(* IEC 61131-3 sources: plc-st-coding-agent/progress/evidence/f14_v3_parallel_20261112/jobs/custom_deepseek-v4pro (part 3) *)

(* ---- self-hard-07.raw_candidate_01.st ---- *)
FUNCTION_BLOCK FB
VAR_INPUT
    mode : INT;
    resetBtn : BOOL;
    scanSeconds : REAL;
    tempSP : REAL;
    tempPV : REAL;
    flowPV : REAL;
    manualFlowSP : REAL;
    manualValve : REAL;
END_VAR
VAR_OUTPUT
    flowSP : REAL;
    valveCommand : REAL;
    fault : BOOL;
    normalMode : BOOL;
END_VAR
VAR
    hasPrev : BOOL := FALSE;
    prevMode : INT := 0;
    prevReset : BOOL := FALSE;
    prevFlowSP : REAL := 0.0;
    prevValveCommand : REAL := 0.0;
    prevET : REAL := 0.0;
    prevEF : REAL := 0.0;
    resetRising : BOOL;
    eT : REAL;
    eF : REAL;
    flowRaw : REAL;
    valveRaw : REAL;
    trialT : REAL;
    trialF : REAL;
END_VAR

fault := (mode < 0) OR (mode > 2) OR (scanSeconds <= 0.0) OR (scanSeconds > 10.0);
resetRising := resetBtn AND NOT prevReset;

IF NOT hasPrev THEN
    normalMode := FALSE;
    flowSP := manualFlowSP;
    valveCommand := manualValve;
ELSIF resetRising THEN
    normalMode := FALSE;
    flowSP := manualFlowSP;
    valveCommand := manualValve;
ELSIF fault THEN
    normalMode := FALSE;
    flowSP := manualFlowSP;
    valveCommand := manualValve;
ELSIF mode <> prevMode THEN
    normalMode := FALSE;
    IF mode = 2 THEN
        flowSP := prevFlowSP;
        valveCommand := prevValveCommand;
    ELSE
        flowSP := manualFlowSP;
        valveCommand := prevValveCommand;
    END_IF;
ELSE
    normalMode := TRUE;
    IF mode = 0 THEN
        flowSP := manualFlowSP;
        valveCommand := manualValve;
    ELSIF mode = 1 THEN
        flowSP := manualFlowSP;
        eF := flowSP - flowPV;
        trialF := prevValveCommand - 2.0 * prevEF + 0.5 * eF * scanSeconds;
        valveRaw := 2.0 * eF + trialF;
        valveCommand := LIMIT(0.0, valveRaw, 100.0);
    ELSIF mode = 2 THEN
        eT := tempSP - tempPV;
        trialT := prevFlowSP - 1.0 * prevET + 0.2 * eT * scanSeconds;
        flowRaw := 1.0 * eT + trialT;
        flowSP := LIMIT(0.0, flowRaw, 50.0);
        eF := flowSP - flowPV;
        trialF := prevValveCommand - 2.0 * prevEF + 0.5 * eF * scanSeconds;
        valveRaw := 2.0 * eF + trialF;
        valveCommand := LIMIT(0.0, valveRaw, 100.0);
    END_IF;
END_IF;

prevFlowSP := flowSP;
prevValveCommand := valveCommand;
prevET := tempSP - tempPV;
prevEF := flowSP - flowPV;
prevMode := mode;
prevReset := resetBtn;
hasPrev := TRUE;

END_FUNCTION_BLOCK

(* ---- self-medium-01.candidate_01.st ---- *)
FUNCTION_BLOCK FB
VAR_INPUT
    recipe : ARRAY[1..8] OF ST_Recipe;   // 配方槽位 1..8，槽位 recipeID=0 表示空
    selSlot : INT;                        // 操作员选中的槽位，合法范围 1..8
    loadCmd : BOOL;                       // 装载命令（上升沿触发一次装载）
    running : BOOL;                       // 当前是否处于生产状态
END_VAR
VAR_OUTPUT
    valid : BOOL;                         // 配方校验通过
    loadedID : INT;                       // 已装载的配方号，无配方时为 0
END_VAR
VAR
    prevLoadCmd  : BOOL;                  // 上一扫描周期的 loadCmd
    prevValid    : BOOL;                  // 上一扫描周期的 valid 输出
    prevLoadedID : INT;                   // 上一扫描周期的 loadedID 输出
    edge         : BOOL;                  // loadCmd 上升沿标志
    slotIndex    : INT;                   // 合法的槽位下标
    slotRecipe   : ST_Recipe;             // 当前选中的配方结构体
    ratioOK      : BOOL;                  // totalRatio 是否在合法区间
    tempOK       : BOOL;                  // temperature 是否在合法区间
END_VAR

    // 计算装载命令的上升沿
    edge := loadCmd AND NOT prevLoadCmd;

    IF running THEN
        // 生产状态：保持上一拍输出，包括刚进入生产的第一拍
        valid := prevValid;
        loadedID := prevLoadedID;
    ELSIF edge THEN
        // 非生产状态且检测到装载命令上升沿
        // 检查槽位是否越界
        IF (selSlot < 1) OR (selSlot > 8) THEN
            // 越界：判为非法，且不得访问数组外内存
            valid := FALSE;
            loadedID := 0;
        ELSE
            // 合法槽位
            slotIndex := selSlot;
            slotRecipe := recipe[slotIndex];

            // 检查槽位是否为空
            IF slotRecipe.recipeID = 0 THEN
                // 空槽：非法
                valid := FALSE;
                loadedID := 0;
            ELSE
                // 检查总配比和温度
                ratioOK := (slotRecipe.totalRatio >= 99.0) AND (slotRecipe.totalRatio <= 101.0);
                tempOK  := (slotRecipe.temperature >= 30.0) AND (slotRecipe.temperature <= 180.0);

                IF ratioOK AND tempOK THEN
                    // 全部校验通过
                    valid := TRUE;
                    loadedID := slotRecipe.recipeID;
                ELSE
                    // 任一校验失败
                    valid := FALSE;
                    loadedID := 0;
                END_IF;
            END_IF;
        END_IF;
    ELSE
        // 无装载沿且未生产：保持上一拍输出
        valid := prevValid;
        loadedID := prevLoadedID;
    END_IF;

    // 更新历史状态
    prevLoadCmd  := loadCmd;
    prevValid    := valid;
    prevLoadedID := loadedID;
END_FUNCTION_BLOCK

(* ---- self-medium-01.candidate_02.st ---- *)
TYPE ST_Recipe :
STRUCT
    recipeID : INT;
    totalRatio : REAL;
    temperature : REAL;
END_STRUCT;
END_TYPE;

FUNCTION_BLOCK FB
VAR_INPUT
    recipe : ARRAY[1..8] OF ST_Recipe;
    selSlot : INT;
    loadCmd : BOOL;
    running : BOOL;
END_VAR
VAR_OUTPUT
    valid : BOOL;
    loadedID : INT;
END_VAR
VAR
    prevLoadCmd  : BOOL;
    prevValid    : BOOL;
    prevLoadedID : INT;
    edge         : BOOL;
    slotIndex    : INT;
    slotRecipe   : ST_Recipe;
    ratioOK      : BOOL;
    tempOK       : BOOL;
END_VAR

    edge := loadCmd AND NOT prevLoadCmd;

    IF running THEN
        (* 生产状态：保持上一拍输出，包括刚进入生产的第一拍 *)
        valid := prevValid;
        loadedID := prevLoadedID;
    ELSIF edge THEN
        (* 非生产状态且检测到装载命令上升沿 *)
        IF (selSlot < 1) OR (selSlot > 8) THEN
            (* 槽位越界：判为非法，不访问数组 *)
            valid := FALSE;
            loadedID := 0;
        ELSE
            slotIndex := selSlot;
            slotRecipe := recipe[slotIndex];

            IF slotRecipe.recipeID = 0 THEN
                (* 空槽：非法 *)
                valid := FALSE;
                loadedID := 0;
            ELSE
                ratioOK := (slotRecipe.totalRatio >= 99.0) AND (slotRecipe.totalRatio <= 101.0);
                tempOK  := (slotRecipe.temperature >= 30.0) AND (slotRecipe.temperature <= 180.0);

                IF ratioOK AND tempOK THEN
                    valid := TRUE;
                    loadedID := slotRecipe.recipeID;
                ELSE
                    valid := FALSE;
                    loadedID := 0;
                END_IF;
            END_IF;
        END_IF;
    ELSE
        (* 无装载沿且未生产：保持上一拍输出 *)
        valid := prevValid;
        loadedID := prevLoadedID;
    END_IF;

    (* 更新历史状态 *)
    prevLoadCmd  := loadCmd;
    prevValid    := valid;
    prevLoadedID := loadedID;
END_FUNCTION_BLOCK

(* ---- self-medium-01.raw_candidate_01.st ---- *)
FUNCTION_BLOCK FB
VAR_INPUT
    recipe : ARRAY[1..8] OF ST_Recipe;   // 配方槽位 1..8，槽位 recipeID=0 表示空
    selSlot : INT;                        // 操作员选中的槽位，合法范围 1..8
    loadCmd : BOOL;                       // 装载命令（上升沿触发一次装载）
    running : BOOL;                       // 当前是否处于生产状态
END_VAR
VAR_OUTPUT
    valid : BOOL;                         // 配方校验通过
    loadedID : INT;                       // 已装载的配方号，无配方时为 0
END_VAR
VAR
    prevLoadCmd  : BOOL;                  // 上一扫描周期的 loadCmd
    prevValid    : BOOL;                  // 上一扫描周期的 valid 输出
    prevLoadedID : INT;                   // 上一扫描周期的 loadedID 输出
    edge         : BOOL;                  // loadCmd 上升沿标志
    slotIndex    : INT;                   // 合法的槽位下标
    slotRecipe   : ST_Recipe;             // 当前选中的配方结构体
    ratioOK      : BOOL;                  // totalRatio 是否在合法区间
    tempOK       : BOOL;                  // temperature 是否在合法区间
END_VAR

    // 计算装载命令的上升沿
    edge := loadCmd AND NOT prevLoadCmd;

    IF running THEN
        // 生产状态：保持上一拍输出，包括刚进入生产的第一拍
        valid := prevValid;
        loadedID := prevLoadedID;
    ELSIF edge THEN
        // 非生产状态且检测到装载命令上升沿
        // 检查槽位是否越界
        IF (selSlot < 1) OR (selSlot > 8) THEN
            // 越界：判为非法，且不得访问数组外内存
            valid := FALSE;
            loadedID := 0;
        ELSE
            // 合法槽位
            slotIndex := selSlot;
            slotRecipe := recipe[slotIndex];

            // 检查槽位是否为空
            IF slotRecipe.recipeID = 0 THEN
                // 空槽：非法
                valid := FALSE;
                loadedID := 0;
            ELSE
                // 检查总配比和温度
                ratioOK := (slotRecipe.totalRatio >= 99.0) AND (slotRecipe.totalRatio <= 101.0);
                tempOK  := (slotRecipe.temperature >= 30.0) AND (slotRecipe.temperature <= 180.0);

                IF ratioOK AND tempOK THEN
                    // 全部校验通过
                    valid := TRUE;
                    loadedID := slotRecipe.recipeID;
                ELSE
                    // 任一校验失败
                    valid := FALSE;
                    loadedID := 0;
                END_IF;
            END_IF;
        END_IF;
    ELSE
        // 无装载沿且未生产：保持上一拍输出
        valid := prevValid;
        loadedID := prevLoadedID;
    END_IF;

    // 更新历史状态
    prevLoadCmd  := loadCmd;
    prevValid    := valid;
    prevLoadedID := loadedID;
END_FUNCTION_BLOCK

(* ---- self-medium-01.raw_candidate_02.st ---- *)
TYPE ST_Recipe :
STRUCT
    recipeID : INT;
    totalRatio : REAL;
    temperature : REAL;
END_STRUCT
END_TYPE

FUNCTION_BLOCK FB
VAR_INPUT
    recipe : ARRAY[1..8] OF ST_Recipe;
    selSlot : INT;
    loadCmd : BOOL;
    running : BOOL;
END_VAR
VAR_OUTPUT
    valid : BOOL;
    loadedID : INT;
END_VAR
VAR
    prevLoadCmd  : BOOL;
    prevValid    : BOOL;
    prevLoadedID : INT;
    edge         : BOOL;
    slotIndex    : INT;
    slotRecipe   : ST_Recipe;
    ratioOK      : BOOL;
    tempOK       : BOOL;
END_VAR

    edge := loadCmd AND NOT prevLoadCmd;

    IF running THEN
        (* 生产状态：保持上一拍输出，包括刚进入生产的第一拍 *)
        valid := prevValid;
        loadedID := prevLoadedID;
    ELSIF edge THEN
        (* 非生产状态且检测到装载命令上升沿 *)
        IF (selSlot < 1) OR (selSlot > 8) THEN
            (* 槽位越界：判为非法，不访问数组 *)
            valid := FALSE;
            loadedID := 0;
        ELSE
            slotIndex := selSlot;
            slotRecipe := recipe[slotIndex];

            IF slotRecipe.recipeID = 0 THEN
                (* 空槽：非法 *)
                valid := FALSE;
                loadedID := 0;
            ELSE
                ratioOK := (slotRecipe.totalRatio >= 99.0) AND (slotRecipe.totalRatio <= 101.0);
                tempOK  := (slotRecipe.temperature >= 30.0) AND (slotRecipe.temperature <= 180.0);

                IF ratioOK AND tempOK THEN
                    valid := TRUE;
                    loadedID := slotRecipe.recipeID;
                ELSE
                    valid := FALSE;
                    loadedID := 0;
                END_IF;
            END_IF;
        END_IF;
    ELSE
        (* 无装载沿且未生产：保持上一拍输出 *)
        valid := prevValid;
        loadedID := prevLoadedID;
    END_IF;

    (* 更新历史状态 *)
    prevLoadCmd  := loadCmd;
    prevValid    := valid;
    prevLoadedID := loadedID;
END_FUNCTION_BLOCK

(* ---- self-medium-02.candidate_01.st ---- *)
FUNCTION_BLOCK FB
VAR_INPUT
    enable : BOOL;
    rawValue : REAL;
END_VAR
VAR_OUTPUT
    filteredValue : REAL;
    windowFull : BOOL;
    sampleCount : INT;
END_VAR
VAR
    buffer : ARRAY[0..7] OF REAL;
    bufIdx : INT := 0;
    cnt : INT := 0;
    sum : REAL;
    i : INT;
END_VAR

IF enable THEN
    buffer[bufIdx] := rawValue;
    bufIdx := bufIdx + 1;
    IF bufIdx >= 8 THEN
        bufIdx := 0;
    END_IF;

    IF cnt < 8 THEN
        cnt := cnt + 1;
    END_IF;

    sum := 0.0;
    FOR i := 0 TO cnt - 1 DO
        sum := sum + buffer[i];
    END_FOR;

    filteredValue := sum / INT_TO_REAL(cnt);
    sampleCount := cnt;
    windowFull := (cnt >= 8);
ELSE
    cnt := 0;
    bufIdx := 0;
    sampleCount := 0;
    windowFull := FALSE;
END_IF;

END_FUNCTION_BLOCK

(* ---- self-medium-02.raw_candidate_01.st ---- *)
FUNCTION_BLOCK FB
VAR_INPUT
    enable : BOOL;
    rawValue : REAL;
END_VAR
VAR_OUTPUT
    filteredValue : REAL;
    windowFull : BOOL;
    sampleCount : INT;
END_VAR
VAR
    buffer : ARRAY[0..7] OF REAL;
    bufIdx : INT := 0;
    cnt : INT := 0;
    sum : REAL;
    i : INT;
END_VAR

IF enable THEN
    buffer[bufIdx] := rawValue;
    bufIdx := bufIdx + 1;
    IF bufIdx >= 8 THEN
        bufIdx := 0;
    END_IF;

    IF cnt < 8 THEN
        cnt := cnt + 1;
    END_IF;

    sum := 0.0;
    FOR i := 0 TO cnt - 1 DO
        sum := sum + buffer[i];
    END_FOR;

    filteredValue := sum / INT_TO_REAL(cnt);
    sampleCount := cnt;
    windowFull := (cnt >= 8);
ELSE
    cnt := 0;
    bufIdx := 0;
    sampleCount := 0;
    windowFull := FALSE;
END_IF;

END_FUNCTION_BLOCK

(* ---- self-medium-03.candidate_01.st ---- *)
FUNCTION_BLOCK FB
VAR_INPUT
    openBtn : BOOL;
    closeBtn : BOOL;
    openLimit : BOOL;
    closeLimit : BOOL;
    obstacle : BOOL;
END_VAR
VAR_OUTPUT
    motorUp : BOOL;
    motorDown : BOOL;
    errorFlag : BOOL;
END_VAR
VAR
    state : INT := 0; (* 0=IDLE, 1=OPENING, 2=CLOSING, 3=FAULT *)
    preOpenBtn : BOOL := FALSE;
    preCloseBtn : BOOL := FALSE;
    risingOpen : BOOL;
    risingClose : BOOL;
    combo : BOOL;
    preCombo : BOOL;
    risingCombo : BOOL;
END_VAR

(* 计算上升沿 *)
risingOpen := openBtn AND NOT preOpenBtn;
risingClose := closeBtn AND NOT preCloseBtn;
combo := openBtn AND closeBtn;
preCombo := preOpenBtn AND preCloseBtn;
risingCombo := combo AND NOT preCombo;

IF obstacle THEN
    (* 障碍优先：任何状态立即停机并置故障 *)
    state := 3;
    motorUp := FALSE;
    motorDown := FALSE;
    errorFlag := TRUE;
ELSE
    IF state = 3 THEN
        (* 无障碍时的故障处理 *)
        IF risingCombo THEN
            (* 双键组合新上升沿：人工复位 *)
            state := 0;
            motorUp := FALSE;
            motorDown := FALSE;
            errorFlag := FALSE;
        ELSE
            (* 保持故障锁存 *)
            motorUp := FALSE;
            motorDown := FALSE;
            errorFlag := TRUE;
        END_IF;
    ELSE
        (* 非故障状态 *)
        IF (state = 1 AND openLimit) OR (state = 2 AND closeLimit) THEN
            (* 到达本方向限位：停机回IDLE *)
            state := 0;
            motorUp := FALSE;
            motorDown := FALSE;
            errorFlag := FALSE;
        ELSE
            IF state = 1 THEN
                (* 开门运行中 *)
                motorUp := TRUE;
                motorDown := FALSE;
                errorFlag := FALSE;
                (* state 保持 1 *)
            ELSIF state = 2 THEN
                (* 关门运行中 *)
                motorUp := FALSE;
                motorDown := TRUE;
                errorFlag := FALSE;
                (* state 保持 2 *)
            ELSE
                (* IDLE状态 *)
                IF risingOpen AND NOT closeBtn AND NOT openLimit THEN
                    state := 1;
                    motorUp := TRUE;
                    motorDown := FALSE;
                    errorFlag := FALSE;
                ELSIF risingClose AND NOT openBtn AND NOT closeLimit THEN
                    state := 2;
                    motorUp := FALSE;
                    motorDown := TRUE;
                    errorFlag := FALSE;
                ELSE
                    motorUp := FALSE;
                    motorDown := FALSE;
                    errorFlag := FALSE;
                    state := 0; (* 保持IDLE *)
                END_IF;
            END_IF;
        END_IF;
    END_IF;
END_IF;

(* 更新上一拍按钮状态 *)
preOpenBtn := openBtn;
preCloseBtn := closeBtn;

END_FUNCTION_BLOCK

(* ---- self-medium-03.raw_candidate_01.st ---- *)
FUNCTION_BLOCK FB
VAR_INPUT
    openBtn : BOOL;
    closeBtn : BOOL;
    openLimit : BOOL;
    closeLimit : BOOL;
    obstacle : BOOL;
END_VAR
VAR_OUTPUT
    motorUp : BOOL;
    motorDown : BOOL;
    errorFlag : BOOL;
END_VAR
VAR
    state : INT := 0; (* 0=IDLE, 1=OPENING, 2=CLOSING, 3=FAULT *)
    preOpenBtn : BOOL := FALSE;
    preCloseBtn : BOOL := FALSE;
    risingOpen : BOOL;
    risingClose : BOOL;
    combo : BOOL;
    preCombo : BOOL;
    risingCombo : BOOL;
END_VAR

(* 计算上升沿 *)
risingOpen := openBtn AND NOT preOpenBtn;
risingClose := closeBtn AND NOT preCloseBtn;
combo := openBtn AND closeBtn;
preCombo := preOpenBtn AND preCloseBtn;
risingCombo := combo AND NOT preCombo;

IF obstacle THEN
    (* 障碍优先：任何状态立即停机并置故障 *)
    state := 3;
    motorUp := FALSE;
    motorDown := FALSE;
    errorFlag := TRUE;
ELSE
    IF state = 3 THEN
        (* 无障碍时的故障处理 *)
        IF risingCombo THEN
            (* 双键组合新上升沿：人工复位 *)
            state := 0;
            motorUp := FALSE;
            motorDown := FALSE;
            errorFlag := FALSE;
        ELSE
            (* 保持故障锁存 *)
            motorUp := FALSE;
            motorDown := FALSE;
            errorFlag := TRUE;
        END_IF
    ELSE
        (* 非故障状态 *)
        IF (state = 1 AND openLimit) OR (state = 2 AND closeLimit) THEN
            (* 到达本方向限位：停机回IDLE *)
            state := 0;
            motorUp := FALSE;
            motorDown := FALSE;
            errorFlag := FALSE;
        ELSE
            IF state = 1 THEN
                (* 开门运行中 *)
                motorUp := TRUE;
                motorDown := FALSE;
                errorFlag := FALSE;
                (* state 保持 1 *)
            ELSIF state = 2 THEN
                (* 关门运行中 *)
                motorUp := FALSE;
                motorDown := TRUE;
                errorFlag := FALSE;
                (* state 保持 2 *)
            ELSE
                (* IDLE状态 *)
                IF risingOpen AND NOT closeBtn AND NOT openLimit THEN
                    state := 1;
                    motorUp := TRUE;
                    motorDown := FALSE;
                    errorFlag := FALSE;
                ELSIF risingClose AND NOT openBtn AND NOT closeLimit THEN
                    state := 2;
                    motorUp := FALSE;
                    motorDown := TRUE;
                    errorFlag := FALSE;
                ELSE
                    motorUp := FALSE;
                    motorDown := FALSE;
                    errorFlag := FALSE;
                    state := 0; (* 保持IDLE *)
                END_IF
            END_IF
        END_IF
    END_IF
END_IF

(* 更新上一拍按钮状态 *)
preOpenBtn := openBtn;
preCloseBtn := closeBtn;

END_FUNCTION_BLOCK

(* ---- self-medium-04.candidate_01.st ---- *)
FUNCTION_BLOCK FB
VAR_INPUT
    startBtn : BOOL;
    resetBtn : BOOL;
    doneSensor : BOOL;
    targetVol : REAL;
    flowVol : REAL;
END_VAR
VAR_OUTPUT
    valveOpen : BOOL;
    fillsToday : INT;
END_VAR
VAR
    prevStart : BOOL := FALSE;
    prevReset : BOOL := FALSE;
    pendingConfirm : BOOL := FALSE;
    accVol : REAL := 0.0;
END_VAR

// 上升沿检测
startRising := startBtn AND NOT prevStart;
resetRising := resetBtn AND NOT prevReset;

IF resetRising THEN
    // 复位优先：清零计数和累计，关阀并清除待确认
    fillsToday := 0;
    accVol := 0.0;
    valveOpen := FALSE;
    pendingConfirm := FALSE;
ELSE
    // 启动处理（空闲或等待确认时）
    IF startRising AND NOT valveOpen THEN
        accVol := 0.0;
        valveOpen := TRUE;
        pendingConfirm := FALSE; // 取消上一瓶待确认
    END_IF;

    // 灌装累加与达标关阀
    IF valveOpen THEN
        accVol := accVol + flowVol;
        IF accVol >= targetVol THEN
            valveOpen := FALSE;
            pendingConfirm := TRUE;
        END_IF;
    END_IF;

    // 确认计数（去抖与饱和处理）
    IF pendingConfirm AND doneSensor THEN
        IF fillsToday < 32767 THEN
            fillsToday := fillsToday + 1;
        END_IF;
        pendingConfirm := FALSE; // 立即清除待确认
    END_IF;
END_IF;

// 更新边沿记忆
prevStart := startBtn;
prevReset := resetBtn;

END_FUNCTION_BLOCK

(* ---- self-medium-04.candidate_02.st ---- *)
FUNCTION_BLOCK FB
VAR_INPUT
    startBtn : BOOL;
    resetBtn : BOOL;
    doneSensor : BOOL;
    targetVol : REAL;
    flowVol : REAL;
END_VAR
VAR_OUTPUT
    valveOpen : BOOL;
    fillsToday : INT;
END_VAR
VAR
    prevStart : BOOL := FALSE;
    prevReset : BOOL := FALSE;
    pendingConfirm : BOOL := FALSE;
    accVol : REAL := 0.0;
    startRising : BOOL;
    resetRising : BOOL;
END_VAR

// 上升沿检测
startRising := startBtn AND NOT prevStart;
resetRising := resetBtn AND NOT prevReset;

IF resetRising THEN
    // 复位优先：清零计数和累计，关阀并清除待确认
    fillsToday := 0;
    accVol := 0.0;
    valveOpen := FALSE;
    pendingConfirm := FALSE;
ELSE
    // 启动处理（空闲或等待确认时）
    IF startRising AND NOT valveOpen THEN
        accVol := 0.0;
        valveOpen := TRUE;
        pendingConfirm := FALSE; // 取消上一瓶待确认
    END_IF;

    // 灌装累加与达标关阀
    IF valveOpen THEN
        accVol := accVol + flowVol;
        IF accVol >= targetVol THEN
            valveOpen := FALSE;
            pendingConfirm := TRUE;
        END_IF;
    END_IF;

    // 确认计数（去抖与饱和处理）
    IF pendingConfirm AND doneSensor THEN
        IF fillsToday < 32767 THEN
            fillsToday := fillsToday + 1;
        END_IF;
        pendingConfirm := FALSE; // 立即清除待确认
    END_IF;
END_IF;

// 更新边沿记忆
prevStart := startBtn;
prevReset := resetBtn;

END_FUNCTION_BLOCK

(* ---- self-medium-04.raw_candidate_01.st ---- *)
FUNCTION_BLOCK FB
VAR_INPUT
    startBtn : BOOL;
    resetBtn : BOOL;
    doneSensor : BOOL;
    targetVol : REAL;
    flowVol : REAL;
END_VAR
VAR_OUTPUT
    valveOpen : BOOL;
    fillsToday : INT;
END_VAR
VAR
    prevStart : BOOL := FALSE;
    prevReset : BOOL := FALSE;
    pendingConfirm : BOOL := FALSE;
    accVol : REAL := 0.0;
END_VAR

// 上升沿检测
startRising := startBtn AND NOT prevStart;
resetRising := resetBtn AND NOT prevReset;

IF resetRising THEN
    // 复位优先：清零计数和累计，关阀并清除待确认
    fillsToday := 0;
    accVol := 0.0;
    valveOpen := FALSE;
    pendingConfirm := FALSE;
ELSE
    // 启动处理（空闲或等待确认时）
    IF startRising AND NOT valveOpen THEN
        accVol := 0.0;
        valveOpen := TRUE;
        pendingConfirm := FALSE; // 取消上一瓶待确认
    END_IF;

    // 灌装累加与达标关阀
    IF valveOpen THEN
        accVol := accVol + flowVol;
        IF accVol >= targetVol THEN
            valveOpen := FALSE;
            pendingConfirm := TRUE;
        END_IF;
    END_IF;

    // 确认计数（去抖与饱和处理）
    IF pendingConfirm AND doneSensor THEN
        IF fillsToday < 32767 THEN
            fillsToday := fillsToday + 1;
        END_IF;
        pendingConfirm := FALSE; // 立即清除待确认
    END_IF;
END_IF;

// 更新边沿记忆
prevStart := startBtn;
prevReset := resetBtn;

END_FUNCTION_BLOCK

(* ---- self-medium-04.raw_candidate_02.st ---- *)
FUNCTION_BLOCK FB
VAR_INPUT
    startBtn : BOOL;
    resetBtn : BOOL;
    doneSensor : BOOL;
    targetVol : REAL;
    flowVol : REAL;
END_VAR
VAR_OUTPUT
    valveOpen : BOOL;
    fillsToday : INT;
END_VAR
VAR
    prevStart : BOOL := FALSE;
    prevReset : BOOL := FALSE;
    pendingConfirm : BOOL := FALSE;
    accVol : REAL := 0.0;
    startRising : BOOL;
    resetRising : BOOL;
END_VAR

// 上升沿检测
startRising := startBtn AND NOT prevStart;
resetRising := resetBtn AND NOT prevReset;

IF resetRising THEN
    // 复位优先：清零计数和累计，关阀并清除待确认
    fillsToday := 0;
    accVol := 0.0;
    valveOpen := FALSE;
    pendingConfirm := FALSE;
ELSE
    // 启动处理（空闲或等待确认时）
    IF startRising AND NOT valveOpen THEN
        accVol := 0.0;
        valveOpen := TRUE;
        pendingConfirm := FALSE; // 取消上一瓶待确认
    END_IF;

    // 灌装累加与达标关阀
    IF valveOpen THEN
        accVol := accVol + flowVol;
        IF accVol >= targetVol THEN
            valveOpen := FALSE;
            pendingConfirm := TRUE;
        END_IF;
    END_IF;

    // 确认计数（去抖与饱和处理）
    IF pendingConfirm AND doneSensor THEN
        IF fillsToday < 32767 THEN
            fillsToday := fillsToday + 1;
        END_IF;
        pendingConfirm := FALSE; // 立即清除待确认
    END_IF;
END_IF;

// 更新边沿记忆
prevStart := startBtn;
prevReset := resetBtn;

END_FUNCTION_BLOCK

(* ---- self-medium-05.candidate_01.st ---- *)
FUNCTION_BLOCK FB
VAR_INPUT
    enable : BOOL;
    resetBtn : BOOL;
    scanSeconds : LREAL;
    steamFlow : LREAL;
    fuelFlow : LREAL;
    steamTemp : LREAL;
    steamPressure : LREAL;
END_VAR
VAR_OUTPUT
    qualified : BOOL;
    dataFault : BOOL;
    qualifiedTon : LREAL;
    fuelTon : LREAL;
    revenue : LREAL;
    cost : LREAL;
    netProfit : LREAL;
END_VAR
VAR
    prevResetBtn : BOOL := FALSE;
    resetRising : BOOL;
END_VAR

    qualified := (steamTemp >= 447.0) AND (steamTemp <= 453.0) AND (steamPressure >= 3750.0) AND (steamPressure <= 3850.0);

    dataFault := (scanSeconds <= 0.0) OR (scanSeconds > 10.0) OR (steamFlow < 0.0) OR (steamFlow > 90.0) OR (fuelFlow < 0.0) OR (fuelFlow > 6.0);

    resetRising := resetBtn AND NOT prevResetBtn;

    IF resetRising THEN
        qualifiedTon := 0.0;
        fuelTon := 0.0;
    ELSE
        IF enable AND NOT dataFault THEN
            fuelTon := fuelTon + (fuelFlow * scanSeconds / 1000.0);
            IF qualified THEN
                qualifiedTon := qualifiedTon + (steamFlow * scanSeconds / 1000.0);
            END_IF;
        END_IF;
    END_IF;

    revenue := qualifiedTon * 280.0;
    cost := fuelTon * 1500.0;
    netProfit := revenue - cost;

    prevResetBtn := resetBtn;

END_FUNCTION_BLOCK

(* ---- self-medium-05.raw_candidate_01.st ---- *)
FUNCTION_BLOCK FB
VAR_INPUT
    enable : BOOL;
    resetBtn : BOOL;
    scanSeconds : LREAL;
    steamFlow : LREAL;
    fuelFlow : LREAL;
    steamTemp : LREAL;
    steamPressure : LREAL;
END_VAR
VAR_OUTPUT
    qualified : BOOL;
    dataFault : BOOL;
    qualifiedTon : LREAL;
    fuelTon : LREAL;
    revenue : LREAL;
    cost : LREAL;
    netProfit : LREAL;
END_VAR
VAR
    prevResetBtn : BOOL := FALSE;
    resetRising : BOOL;
END_VAR

    qualified := (steamTemp >= 447.0) AND (steamTemp <= 453.0) AND (steamPressure >= 3750.0) AND (steamPressure <= 3850.0);

    dataFault := (scanSeconds <= 0.0) OR (scanSeconds > 10.0) OR (steamFlow < 0.0) OR (steamFlow > 90.0) OR (fuelFlow < 0.0) OR (fuelFlow > 6.0);

    resetRising := resetBtn AND NOT prevResetBtn;

    IF resetRising THEN
        qualifiedTon := 0.0;
        fuelTon := 0.0;
    ELSE
        IF enable AND NOT dataFault THEN
            fuelTon := fuelTon + (fuelFlow * scanSeconds / 1000.0);
            IF qualified THEN
                qualifiedTon := qualifiedTon + (steamFlow * scanSeconds / 1000.0);
            END_IF;
        END_IF;
    END_IF;

    revenue := qualifiedTon * 280.0;
    cost := fuelTon * 1500.0;
    netProfit := revenue - cost;

    prevResetBtn := resetBtn;

END_FUNCTION_BLOCK

(* ---- self-medium-06.candidate_01.st ---- *)
FUNCTION_BLOCK FB
VAR_INPUT
    enable : BOOL;
    resetBtn : BOOL;
    sensorValid : BOOL;
    setpoint : REAL;
    temperature : REAL;
    scanSeconds : REAL;
    bias : REAL;
END_VAR
VAR_OUTPUT
    power : REAL;
    correction : REAL;
    fault : BOOL;
END_VAR
VAR
    ePrev : REAL := 0.0;
    historyValid : BOOL := FALSE;
    prevResetBtn : BOOL := FALSE;
    e : REAL;
    de : REAL;
    x : REAL;
    y : REAL;
    muN_x : REAL;
    muZ_x : REAL;
    muP_x : REAL;
    muN_y : REAL;
    muZ_y : REAL;
    muP_y : REAL;
    sumW : REAL;
    sumWC : REAL;
    risingReset : BOOL;
END_VAR

fault := NOT sensorValid OR (scanSeconds <= 0.0) OR (scanSeconds > 10.0);
risingReset := resetBtn AND NOT prevResetBtn;
e := setpoint - temperature;

IF (NOT enable) OR fault OR risingReset THEN
    power := 0.0;
    correction := 0.0;
    ePrev := 0.0;
    historyValid := FALSE;
ELSE
    IF historyValid THEN
        de := (e - ePrev) / scanSeconds;
    ELSE
        de := 0.0;
    END_IF;

    x := e / 10.0;
    IF x < -1.0 THEN
        x := -1.0;
    ELSIF x > 1.0 THEN
        x := 1.0;
    END_IF;

    y := de / 2.0;
    IF y < -1.0 THEN
        y := -1.0;
    ELSIF y > 1.0 THEN
        y := 1.0;
    END_IF;

    muN_x := MAX(-x, 0.0);
    muZ_x := 1.0 - ABS(x);
    muP_x := MAX(x, 0.0);

    muN_y := MAX(-y, 0.0);
    muZ_y := 1.0 - ABS(y);
    muP_y := MAX(y, 0.0);

    sumW := (muN_x * muN_y) + (muN_x * muZ_y) + (muN_x * muP_y)
          + (muZ_x * muN_y) + (muZ_x * muZ_y) + (muZ_x * muP_y)
          + (muP_x * muN_y) + (muP_x * muZ_y) + (muP_x * muP_y);

    sumWC := (muN_x * muN_y * (-30.0)) + (muN_x * muZ_y * (-20.0)) + (muN_x * muP_y * (-10.0))
           + (muZ_x * muN_y * (-10.0)) + (muZ_x * muZ_y * 0.0) + (muZ_x * muP_y * 10.0)
           + (muP_x * muN_y * 10.0) + (muP_x * muZ_y * 20.0) + (muP_x * muP_y * 30.0);

    IF sumW = 0.0 THEN
        correction := 0.0;
    ELSE
        correction := sumWC / sumW;
    END_IF;

    power := LIMIT(0.0, bias + correction, 100.0);

    ePrev := e;
    historyValid := TRUE;
END_IF;

prevResetBtn := resetBtn;

END_FUNCTION_BLOCK

(* ---- self-medium-06.raw_candidate_01.st ---- *)
FUNCTION_BLOCK FB
VAR_INPUT
    enable : BOOL;
    resetBtn : BOOL;
    sensorValid : BOOL;
    setpoint : REAL;
    temperature : REAL;
    scanSeconds : REAL;
    bias : REAL;
END_VAR
VAR_OUTPUT
    power : REAL;
    correction : REAL;
    fault : BOOL;
END_VAR
VAR
    ePrev : REAL := 0.0;
    historyValid : BOOL := FALSE;
    prevResetBtn : BOOL := FALSE;
    e : REAL;
    de : REAL;
    x : REAL;
    y : REAL;
    muN_x : REAL;
    muZ_x : REAL;
    muP_x : REAL;
    muN_y : REAL;
    muZ_y : REAL;
    muP_y : REAL;
    sumW : REAL;
    sumWC : REAL;
    risingReset : BOOL;
END_VAR

fault := NOT sensorValid OR (scanSeconds <= 0.0) OR (scanSeconds > 10.0);
risingReset := resetBtn AND NOT prevResetBtn;
e := setpoint - temperature;

IF (NOT enable) OR fault OR risingReset THEN
    power := 0.0;
    correction := 0.0;
    ePrev := 0.0;
    historyValid := FALSE;
ELSE
    IF historyValid THEN
        de := (e - ePrev) / scanSeconds;
    ELSE
        de := 0.0;
    END_IF;

    x := e / 10.0;
    IF x < -1.0 THEN
        x := -1.0;
    ELSIF x > 1.0 THEN
        x := 1.0;
    END_IF;

    y := de / 2.0;
    IF y < -1.0 THEN
        y := -1.0;
    ELSIF y > 1.0 THEN
        y := 1.0;
    END_IF;

    muN_x := MAX(-x, 0.0);
    muZ_x := 1.0 - ABS(x);
    muP_x := MAX(x, 0.0);

    muN_y := MAX(-y, 0.0);
    muZ_y := 1.0 - ABS(y);
    muP_y := MAX(y, 0.0);

    sumW := (muN_x * muN_y) + (muN_x * muZ_y) + (muN_x * muP_y)
          + (muZ_x * muN_y) + (muZ_x * muZ_y) + (muZ_x * muP_y)
          + (muP_x * muN_y) + (muP_x * muZ_y) + (muP_x * muP_y);

    sumWC := (muN_x * muN_y * (-30.0)) + (muN_x * muZ_y * (-20.0)) + (muN_x * muP_y * (-10.0))
           + (muZ_x * muN_y * (-10.0)) + (muZ_x * muZ_y * 0.0) + (muZ_x * muP_y * 10.0)
           + (muP_x * muN_y * 10.0) + (muP_x * muZ_y * 20.0) + (muP_x * muP_y * 30.0);

    IF sumW = 0.0 THEN
        correction := 0.0;
    ELSE
        correction := sumWC / sumW;
    END_IF;

    power := LIMIT(0.0, bias + correction, 100.0);

    ePrev := e;
    historyValid := TRUE;
END_IF;

prevResetBtn := resetBtn;

END_FUNCTION_BLOCK
